(* IEC 61131-3 sources: volt/packages/volt-lsp-iec/test-corpus/pro2193/Device/Plc Logic/Application/09 Misc/Library Manager/SysFile, 24 files *)

(* ---- ACCESS_MODE.dut ---- *)
TYPE ACCESS_MODE :
(
	AM_READ,
	AM_WRITE,
	AM_APPEND,
	AM_READ_PLUS,
	AM_WRITE_PLUS,
	AM_APPEND_PLUS
);
END_TYPE

(* ---- SYS_FILE_STATUS.dut ---- *)
TYPE SYS_FILE_STATUS :
(
	FS_OK,
	FS_NO_FILE,
	FS_ILLEGAL_POS,
	FS_FULL,
	FS_EOF
);
END_TYPE

(* ---- SYS_FILETIME.dut ---- *)
TYPE SYS_FILETIME :
STRUCT
	TCREATION : UDINT;
	TLASTACCESS : UDINT;
	TLASTMODIFICATION : UDINT;
END_STRUCT
END_TYPE

(* ---- SYSFILECLOSE.pou ---- *)
FUNCTION SYSFILECLOSE : RTS_IEC_RESULT
VAR_INPUT
	HFILE : RTS_IEC_HANDLE;
END_VAR
END_FUNCTION

(* ---- SYSFILECOPY.pou ---- *)
FUNCTION SYSFILECOPY : RTS_IEC_RESULT
VAR_INPUT
	SZDESTFILENAME : REFERENCE TO STRING;
	SZSOURCEFILENAME : REFERENCE TO STRING;
	PULCOPIED : POINTER TO __XWORD;
END_VAR
END_FUNCTION

(* ---- SYSFILEDELETE.pou ---- *)
FUNCTION SYSFILEDELETE : RTS_IEC_RESULT
VAR_INPUT
	SZFILENAME : REFERENCE TO STRING;
END_VAR
END_FUNCTION

(* ---- SYSFILEDELETEBYHANDLE.pou ---- *)
FUNCTION SYSFILEDELETEBYHANDLE : RTS_IEC_RESULT
VAR_INPUT
	HFILE : RTS_IEC_HANDLE;
END_VAR
END_FUNCTION

(* ---- SYSFILEEOF.pou ---- *)
FUNCTION SYSFILEEOF : RTS_IEC_RESULT
VAR_INPUT
	HFILE : RTS_IEC_HANDLE;
END_VAR
END_FUNCTION

(* ---- SYSFILEFLUSH.pou ---- *)
FUNCTION SYSFILEFLUSH : RTS_IEC_RESULT
VAR_INPUT
	HFILE : RTS_IEC_HANDLE;
END_VAR
END_FUNCTION

(* ---- SYSFILEGETNAME.pou ---- *)
FUNCTION SYSFILEGETNAME : POINTER TO STRING
VAR_INPUT
	HFILE : RTS_IEC_HANDLE;
END_VAR
END_FUNCTION

(* ---- SYSFILEGETNAME2.pou ---- *)
FUNCTION SYSFILEGETNAME2 : POINTER TO STRING
VAR_INPUT
	HFILE : RTS_IEC_HANDLE;
	PRESULT : POINTER TO RTS_IEC_RESULT;
END_VAR
END_FUNCTION

(* ---- SYSFILEGETPATH.pou ---- *)
FUNCTION SYSFILEGETPATH : RTS_IEC_RESULT
VAR_INPUT
	SZFILENAME : REFERENCE TO STRING;
	DIMAXLEN : DINT;
END_VAR
VAR_IN_OUT
	SZPATH : STRING;
END_VAR
END_FUNCTION

(* ---- SYSFILEGETPOS.pou ---- *)
FUNCTION SYSFILEGETPOS : RTS_IEC_RESULT
VAR_INPUT
	HFILE : RTS_IEC_HANDLE;
	PULPOS : POINTER TO __XWORD;
END_VAR
END_FUNCTION

(* ---- SYSFILEGETSIZE.pou ---- *)
FUNCTION SYSFILEGETSIZE : __XWORD
VAR_INPUT
	SZFILENAME : REFERENCE TO STRING;
	PRESULT : POINTER TO RTS_IEC_RESULT;
END_VAR
END_FUNCTION

(* ---- SYSFILEGETSIZEBYHANDLE.pou ---- *)
FUNCTION SYSFILEGETSIZEBYHANDLE : __XWORD
VAR_INPUT
	HFILE : RTS_IEC_HANDLE;
	PRESULT : POINTER TO RTS_IEC_RESULT;
END_VAR
END_FUNCTION

(* ---- SYSFILEGETSTATUS.pou ---- *)
FUNCTION SYSFILEGETSTATUS : SYS_FILE_STATUS
VAR_INPUT
	HFILE : RTS_IEC_HANDLE;
END_VAR
END_FUNCTION

(* ---- SYSFILEGETSTATUS2.pou ---- *)
FUNCTION SYSFILEGETSTATUS2 : SYS_FILE_STATUS
VAR_INPUT
	HFILE : RTS_IEC_HANDLE;
	PRESULT : POINTER TO RTS_IEC_RESULT;
END_VAR
END_FUNCTION

(* ---- SYSFILEGETTIME.pou ---- *)
FUNCTION SYSFILEGETTIME : RTS_IEC_RESULT
VAR_INPUT
	SZFILENAME : REFERENCE TO STRING;
	PTFILETIME : POINTER TO SYS_FILETIME;
END_VAR
END_FUNCTION

(* ---- SYSFILEOPEN.pou ---- *)
FUNCTION SYSFILEOPEN : RTS_IEC_HANDLE
VAR_INPUT
	SZFILE : REFERENCE TO STRING;
	AM : ACCESS_MODE;
	PRESULT : POINTER TO RTS_IEC_RESULT;
END_VAR
END_FUNCTION

(* ---- SYSFILEREAD.pou ---- *)
FUNCTION SYSFILEREAD : __XWORD
VAR_INPUT
	HFILE : RTS_IEC_HANDLE;
	PBYBUFFER : POINTER TO BYTE;
	ULSIZE : __XWORD;
	PRESULT : POINTER TO RTS_IEC_RESULT;
END_VAR
END_FUNCTION

(* ---- SYSFILERENAME.pou ---- *)
FUNCTION SYSFILERENAME : RTS_IEC_RESULT
VAR_INPUT
	SZOLDFILENAME : REFERENCE TO STRING;
	SZNEWFILENAME : REFERENCE TO STRING;
END_VAR
END_FUNCTION

(* ---- SYSFILESETPOS.pou ---- *)
FUNCTION SYSFILESETPOS : RTS_IEC_RESULT
VAR_INPUT
	HFILE : RTS_IEC_HANDLE;
	ULOFFSET : __XWORD;
END_VAR
END_FUNCTION

(* ---- SYSFILETRUNCATE.pou ---- *)
FUNCTION SYSFILETRUNCATE : RTS_IEC_RESULT
VAR_INPUT
	HFILE : RTS_IEC_HANDLE;
	ULSIZENEW : __XWORD;
END_VAR
END_FUNCTION

(* ---- SYSFILEWRITE.pou ---- *)
FUNCTION SYSFILEWRITE : __XWORD
VAR_INPUT
	HFILE : RTS_IEC_HANDLE;
	PBYBUFFER : POINTER TO BYTE;
	ULSIZE : __XWORD;
	PRESULT : POINTER TO RTS_IEC_RESULT;
END_VAR
END_FUNCTION
